Fanuc KAREL source: kb00078.KL

-- PROVISIONAL review KL for V940-1; original PC SHA256 984243dbf848b7af47dab3e417f29e9acd5010d13b9ddebb547e7182d5dac268
-- Incomplete behavior may be omitted. Consult companion uncertainty JSON. Do not deploy.
PROGRAM KB00078
%NOLOCKGROUP
BEGIN
  -- V9_ZERO_TABLE_METADATA_HINT layout=0002_ascii; no indexed target words; source/name/runtime held
  -- UNRESOLVED_PC offsets 5-21; opcodes 27,22,31,23
  -- UNRESOLVED_PC offsets 26-30; opcodes 7F
END KB00078
